// TIA Portal V21 export
// export: Created 2026-11-21T13:24:04.8975165Z, ExportSetting WithDefaults, DisplayName Totally Integrated Automation Portal, DisplayVersion V21, DisplayName STEP 7 Professional, DisplayVersion V21, DisplayName STEP 7 Safety, DisplayVersion V21, DisplayName Tech WebApplication, DisplayVersion V21, DisplayName WinCC Basic/Comfort/Advanced, DisplayVersion V21, DisplayName WinCC Unified, DisplayVersion V21
VAR_GLOBAL   // PLC tag table "Safety IO"
   FI_Start AT %I0.0 : Bool;   // Start button, fail-safe input
   FI_Stop AT %I0.1 : Bool;   // Stop button, fail-safe input
   FI_DoorClosed AT %I0.2 : Bool;   // Door switch
   FI_GuardClosed AT %I20.0 : Bool;   // Guard door switch on the remote station
   FQ_Motor AT %Q10.0 : Bool;   // Motor contactor, fail-safe output
   FQ_Lamp AT %Q10.1 : Bool;   // Signal lamp, fail-safe output
END_VAR
